{attribute 'qualified_only'}
VAR_GLOBAL CONSTANT
    UNIT_STATE_TIMEOUT_DEFAULT : TIME := T#10S;
END_VAR
VAR_GLOBAL
END_VAR

(* stored: Version 1.1.0.1, ProductVersion 3.1.4024.16
   GVL GVL_PackML: Id {2947b172-aaeb-4f48-90df-804d53a6e375} *)
